FUNCTION_BLOCK VacuumDriver (* Composite Function Block Type *)
  (* Standard: 61499-2 *)
  (* Version 0.0, 7/2/2026, template *)
  PACKAGE Main;
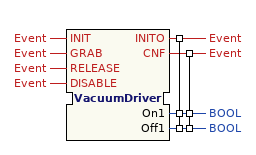
  EVENT_INPUT
    INIT; (* Initialization Request *)
    GRAB; (* Normal Execution Request *)
    RELEASE;
    DISABLE;
  END_EVENT
  EVENT_OUTPUT
    INITO WITH On1, Off1; (* Initialization Confirm *)
    CNF WITH On1, Off1; (* Execution Confirmation *)
  END_EVENT
  VAR_OUTPUT
    On1 : BOOL; (* Output event qualifier *)
    Off1 : BOOL;
  END_VAR
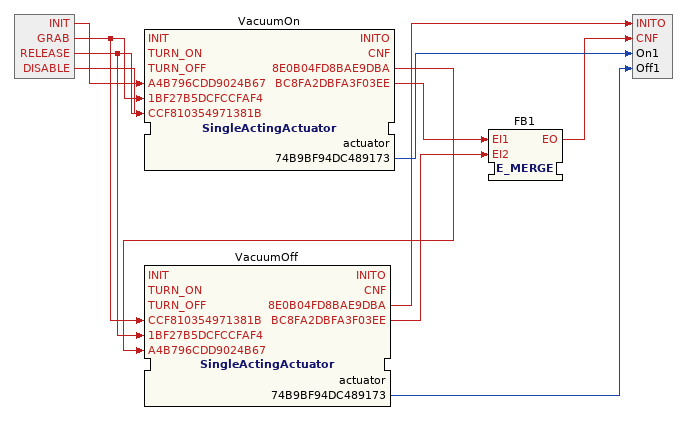
  FBS
    VacuumOn : SingleActingActuator;
    VacuumOff : SingleActingActuator;
    FB1 : E_MERGE;
  END_FBS
  EVENT_CONNECTIONS
    INIT TO VacuumOn.A4B796CDD9024B67;
    FB1.EO TO CNF;
    VacuumOff.8E0B04FD8BAE9DBA TO INITO;
    GRAB TO VacuumOff.CCF810354971381B;
    RELEASE TO VacuumOff.1BF27B5DCFCCFAF4;
    GRAB TO VacuumOn.1BF27B5DCFCCFAF4;
    RELEASE TO VacuumOn.CCF810354971381B;
    DISABLE TO VacuumOn.CCF810354971381B;
    VacuumOn.8E0B04FD8BAE9DBA TO VacuumOff.A4B796CDD9024B67;
    VacuumOn.BC8FA2DBFA3F03EE TO FB1.EI1;
    VacuumOff.BC8FA2DBFA3F03EE TO FB1.EI2;
  END_CONNECTIONS
  DATA_CONNECTIONS
    VacuumOff.74B9BF94DC489173 TO Off1;
    VacuumOn.74B9BF94DC489173 TO On1;
  END_CONNECTIONS
END_FUNCTION_BLOCK
